(* Logix 5000 project; controller SmartManufacturingCell Emulate 5570 rev 33.11; software revision 33.03; part 4 of 5 *)
(* tags used below, declared in another part *)
   Production_CycleHealthy : BOOL;
   SequenceAtScan : DINT;
   StatisticsResetAccepted : BOOL;
   StatisticsResetONS : BOOL;
   Stats_ExitElapsed : REAL;
   Stats_HasPreviousExit : BOOL;
   Stats_RateElapsed : REAL;
   Stats_WindowCount : DINT;
   Conveyor_Flt_FailToStart : BOOL;   // Conveyor commanded but running feedback missing for 2 s Latched; clear cell, remove cause, then fresh Reset.
   Exit_Flt_DischargeTimeout : BOOL;   // Good or reject bottle departure not confirmed within 3 s Latched; clear cell, remove cause, then fresh Reset.
   Exit_Sts_GoodCompletePulse : BOOL;   // Exit Sts GoodCompletePulse
   Exit_Sts_RejectCompletePulse : BOOL;   // Exit Sts RejectCompletePulse
   Exit_Sts_State : DINT;   // 0 Empty; 10 Waiting; 20 Good discharge; 30 Extending; 40 Reject discharge; 50 Retracting; 60 Complete; 90 Faulted
   Filling_Flt_FillTimeout : BOOL;   // Fill completion not received within 4 s Latched; clear cell, remove cause, then fresh Reset.
   Filling_Flt_ValveFailToClose : BOOL;   // Fill valve did not close within 2 s Latched; clear cell, remove cause, then fresh Reset.
   Filling_Sts_ActiveFillTimeMs : DINT;   // Sampled fill duration for current bottle
   HMI_Cmd_Acknowledge : BOOL;   // Acknowledge alarm indication; does not reset faults
   HMI_Cmd_ClearCell : BOOL;   // Request removal of simulated bottles during fault recovery
   HMI_Cmd_ResetStatistics : BOOL;   // Clear production statistics only when Stopped and cell empty
   HMI_Cmd_Start : BOOL;   // Request automatic production start
   HMI_Cmd_Stop : BOOL;   // Request controlled production stop
   HMI_Sim_BottleMissingAtFill : BOOL;   // Suppress Fill photoeye while retaining simulated bottle presence. Simulation test only.
   HMI_Sim_ConveyorFailToStart : BOOL;   // Suppress conveyor running feedback. Simulation test only.
   HMI_Sim_FillFailToComplete : BOOL;   // Suppress simulated filling completion. Simulation test only.
   HMI_Sim_FillValveFailToClose : BOOL;   // Suppress fill valve closed feedback. Simulation test only.
   HMI_Sim_GoodDischargeJam : BOOL;   // Prevent good bottle departure. Simulation test only.
   HMI_Sim_IndexJam : BOOL;   // Prevent simulated index travel from completing. Simulation test only.
   HMI_Sim_IndexPositionMismatch : BOOL;   // Invert simulated Fill occupancy on transfer to test confirmation. Simulation test only.
   HMI_Sim_RejectDischargeJam : BOOL;   // Prevent rejected bottle departure. Simulation test only.
   HMI_Sim_RejectFailToExtend : BOOL;   // Suppress reject extended feedback. Simulation test only.
   HMI_Sim_RejectFailToRetract : BOOL;   // Suppress reject retracted feedback. Simulation test only.
   Inspection_Flt_Timeout : BOOL;   // Inspection did not finish within 3 s Latched; clear cell, remove cause, then fresh Reset.
   Production_Bottles : UDT_Bottle[4];
   Production_Flt_IndexConfirmTimeout : BOOL;   // Post-index positions not confirmed within 1 s Latched; clear cell, remove cause, then fresh Reset.
   Production_Flt_IndexInterlock : BOOL;   // Movement interlock lost during indexing Latched; clear cell, remove cause, then fresh Reset.
   Production_Flt_IndexTimeout : BOOL;   // Index completion not received within 3 s Latched; clear cell, remove cause, then fresh Reset.
   Production_Flt_InvalidConfiguration : BOOL;   // Fill or inspection time outside permitted limits Latched; clear cell, remove cause, then fresh Reset.
   Production_Flt_InvalidState : BOOL;   // Machine, sequence, station state, or mode combination invalid Latched; clear cell, remove cause, then fresh Reset.
   Production_Flt_StartupRecoveryRequired : BOOL;   // Restart found bottles or interrupted activity Latched; clear cell, remove cause, then fresh Reset.
   Production_Flt_TrackingMismatch : BOOL;   // Stationary bottle tracking and sensors disagree or processing history invalid Latched; clear cell, remove cause, then fr
   Production_Stats_FaultSeconds : REAL;   // FaultSeconds based on 20 ms scheduled executions; not a wall-clock historian.
   Production_Stats_GoodCount : DINT;   // Retained GoodCount; count only confirmed departures (recovery losses separate).
   Production_Stats_LastCycleSeconds : REAL;   // LastCycleSeconds based on 20 ms scheduled executions; not a wall-clock historian.
   Production_Stats_RatePerMinute : REAL;   // RatePerMinute based on 20 ms scheduled executions; not a wall-clock historian.
   Production_Stats_RecoveryLossCount : DINT;   // Retained RecoveryLossCount; count only confirmed departures (recovery losses separate).
   Production_Stats_RejectCount : DINT;   // Retained RejectCount; count only confirmed departures (recovery losses separate).
   Production_Stats_RunSeconds : REAL;   // RunSeconds based on 20 ms scheduled executions; not a wall-clock historian.
   Production_Stats_StoppedSeconds : REAL;   // StoppedSeconds based on 20 ms scheduled executions; not a wall-clock historian.
   Production_Stats_TotalCount : DINT;   // Retained TotalCount; count only confirmed departures (recovery losses separate).
   Production_Sts_ClearCellAccepted : BOOL;
   Production_Sts_CounterSaturated : BOOL;   // Production Sts CounterSaturated
   Production_Sts_IndexAllowed : BOOL;
   Production_Sts_IndexCommitted : BOOL;   // Bottle records transferred for the current confirmed index; cleared outside ConfirmPositions.
   Production_Sts_LoadAccepted : BOOL;
   Production_Sts_SequenceState : DINT;   // 0 = Idle 10 = ProcessStations 20 = Indexing 30 = ConfirmPositions
   Reject_Flt_FailToExtend : BOOL;   // Reject actuator did not extend within 2 s Latched; clear cell, remove cause, then fresh Reset.
   Reject_Flt_FailToRetract : BOOL;   // Reject actuator did not retract within 2 s Latched; clear cell, remove cause, then fresh Reset.
   Sim_In_ConveyorRunning : BOOL;   // Simulated conveyor movement feedback
   Sim_In_EntryPE : BOOL;   // Simulated bottle detected at entry
   Sim_In_ExitPE : BOOL;   // Simulated bottle detected at Reject/Exit position
   Sim_In_FillComplete : BOOL;   // Sim In FillComplete
   Sim_In_FillPE : BOOL;   // Simulated bottle detected at filling position
   Sim_In_FillValveClosed : BOOL;   // Simulated fill valve confirmed closed
   Sim_In_GoodExitPE : BOOL;   // Bottle detected passing through good discharge path
   Sim_In_IndexComplete : BOOL;   // Simulated conveyor completed one station-spacing movement
   Sim_In_InspectionPE : BOOL;   // Simulated bottle detected at inspection position
   Sim_In_RejectExitPE : BOOL;   // Bottle detected passing through reject discharge path
   Sim_In_RejectExtended : BOOL;   // Simulated reject actuator confirmed extended
   Sim_In_RejectRetracted : BOOL;   // Simulated reject actuator confirmed retracted
   Sim_Out_ConveyorRun : BOOL;   // Command simulated conveyor to run
   Sim_Out_FillValveOpen : BOOL;   // Command simulated fill valve to open
   Sim_Out_GoodDischargeRun : BOOL;   // Command simulated good-bottle discharge mechanism to run
   Sim_Out_RejectExtend : BOOL;   // Command simulated reject actuator to extend
   Sim_Sts_BottlesPresent : BOOL;   // Sim Sts BottlesPresent
   Sys_Sts_ActiveAlarmCount : DINT;   // Number of active latched faults
   Sys_Sts_AlarmUnacknowledged : BOOL;   // Sys Sts AlarmUnacknowledged
   Sys_Sts_AutoMode : BOOL;   // Auto mode accepted and active
   Sys_Sts_CellEmpty : BOOL;   // Sys Sts CellEmpty
   Sys_Sts_EquipmentHome : BOOL;   // Sys Sts EquipmentHome
   Sys_Sts_FirstFaultCode : DINT;   // Lowest active fault code; zero means none
   Sys_Sts_MachineState : DINT;   // 0 = Stopped 10 = Running 20 = Stopping 30 = Faulted
   Sys_Sts_ManualMode : BOOL;   // Manual mode accepted and active
   Sys_Sts_StartupReady : BOOL;   // Sys Sts StartupReady
(* Program_Production, continued *)

ROUTINE Production_Sequence   (* ladder *)
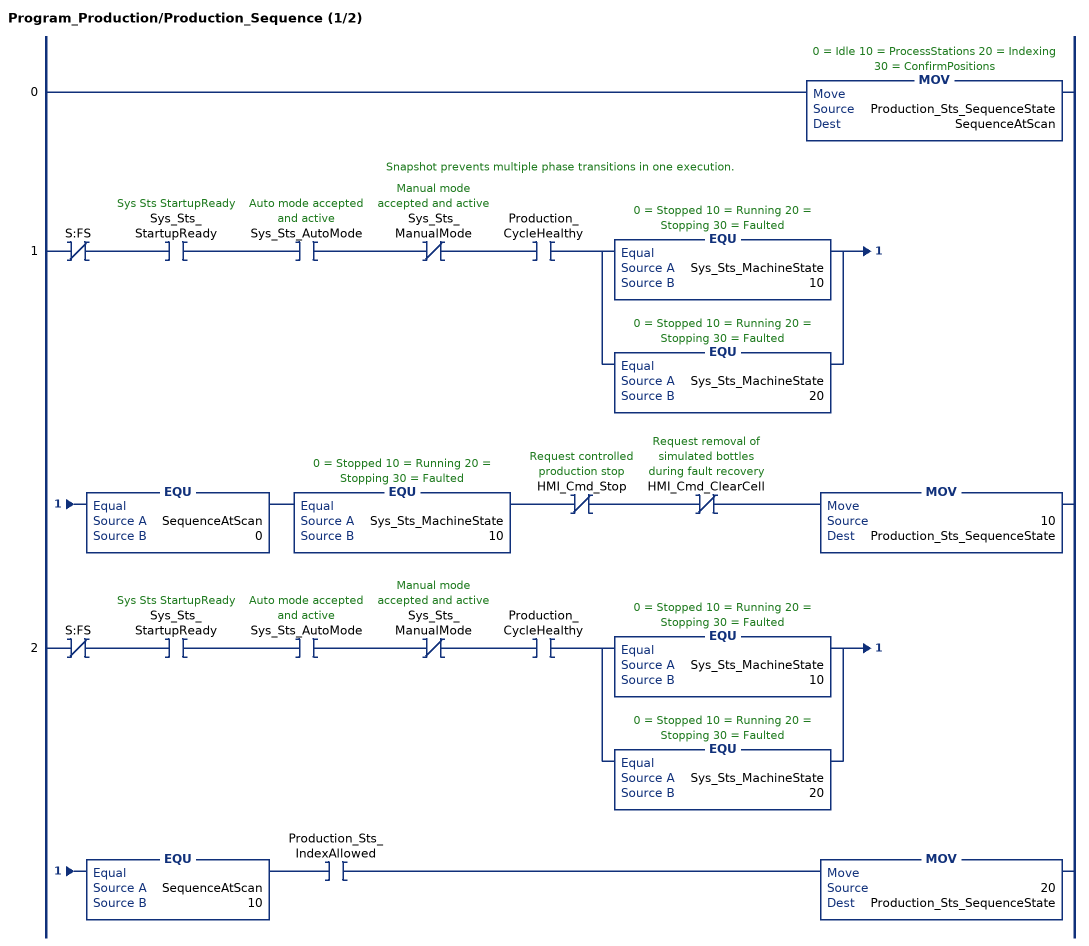
   0: MOV(Production_Sts_SequenceState,SequenceAtScan);
   // Snapshot prevents multiple phase transitions in one execution.
   1: XIO(S:FS)XIC(Sys_Sts_StartupReady)XIC(Sys_Sts_AutoMode)XIO(Sys_Sts_ManualMode)XIC(Production_CycleHealthy)[EQU(Sys_Sts_MachineState,10) ,EQU(Sys_Sts_MachineState,20) ]EQU(SequenceAtScan,0)EQU(Sys_Sts_MachineState,10)XIO(HMI_Cmd_Stop)XIO(HMI_Cmd_ClearCell)MOV(10,Production_Sts_SequenceState);
   2: XIO(S:FS)XIC(Sys_Sts_StartupReady)XIC(Sys_Sts_AutoMode)XIO(Sys_Sts_ManualMode)XIC(Production_CycleHealthy)[EQU(Sys_Sts_MachineState,10) ,EQU(Sys_Sts_MachineState,20) ]EQU(SequenceAtScan,10)XIC(Production_Sts_IndexAllowed)MOV(20,Production_Sts_SequenceState);
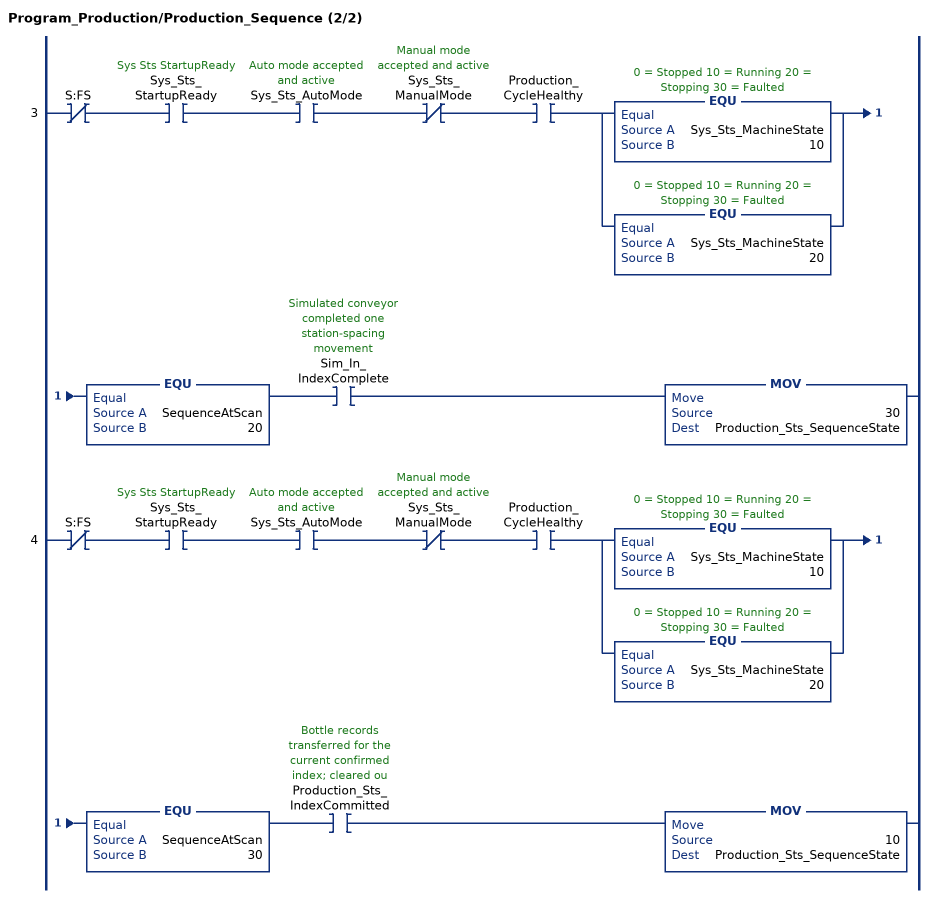
   3: XIO(S:FS)XIC(Sys_Sts_StartupReady)XIC(Sys_Sts_AutoMode)XIO(Sys_Sts_ManualMode)XIC(Production_CycleHealthy)[EQU(Sys_Sts_MachineState,10) ,EQU(Sys_Sts_MachineState,20) ]EQU(SequenceAtScan,20)XIC(Sim_In_IndexComplete)MOV(30,Production_Sts_SequenceState);
   4: XIO(S:FS)XIC(Sys_Sts_StartupReady)XIC(Sys_Sts_AutoMode)XIO(Sys_Sts_ManualMode)XIC(Production_CycleHealthy)[EQU(Sys_Sts_MachineState,10) ,EQU(Sys_Sts_MachineState,20) ]EQU(SequenceAtScan,30)XIC(Production_Sts_IndexCommitted)MOV(10,Production_Sts_SequenceState);
END_ROUTINE

ROUTINE Production_Statistics   (* structured text *)
   // One event per confirmed departure. Recovery clear losses are counted separately.
   IF Exit_Sts_GoodCompletePulse OR Exit_Sts_RejectCompletePulse THEN
       IF Production_Stats_TotalCount < 2147483647 THEN
           Production_Stats_TotalCount := Production_Stats_TotalCount + 1;
           IF Exit_Sts_GoodCompletePulse THEN
               Production_Stats_GoodCount := Production_Stats_GoodCount + 1;
           ELSE
               Production_Stats_RejectCount := Production_Stats_RejectCount + 1;
           END_IF;
       ELSE
           Production_Sts_CounterSaturated := 1;
       END_IF;
       IF Stats_HasPreviousExit THEN
           Production_Stats_LastCycleSeconds := Stats_ExitElapsed;
       END_IF;
       Stats_HasPreviousExit := 1;
       Stats_ExitElapsed := 0.0;
       Stats_WindowCount := Stats_WindowCount + 1;
       Production_Bottles[3].Occupied := 0;
       Production_Bottles[3].FillComplete := 0;
       Production_Bottles[3].InspectionComplete := 0;
       Production_Bottles[3].RejectRequired := 0;
   END_IF;
   IF (Sys_Sts_MachineState = 10) OR (Sys_Sts_MachineState = 20) THEN
       Production_Stats_RunSeconds := Production_Stats_RunSeconds + 0.02;
       Stats_ExitElapsed := Stats_ExitElapsed + 0.02;
   ELSIF Sys_Sts_MachineState = 30 THEN
       Production_Stats_FaultSeconds := Production_Stats_FaultSeconds + 0.02;
   ELSE
       Production_Stats_StoppedSeconds := Production_Stats_StoppedSeconds + 0.02;
   END_IF;
   Stats_RateElapsed := Stats_RateElapsed + 0.02;
   IF Stats_RateElapsed >= 60.0 THEN
       Production_Stats_RatePerMinute := Stats_WindowCount * 60.0 / Stats_RateElapsed;
       Stats_RateElapsed := 0.0;
       Stats_WindowCount := 0;
   END_IF;
   IF S:FS THEN
       Stats_ExitElapsed := 0.0;
       Stats_HasPreviousExit := 0;
       Stats_RateElapsed := 0.0;
       Stats_WindowCount := 0;
       Production_Stats_RatePerMinute := 0.0;
   END_IF;
   IF StatisticsResetAccepted THEN
       Production_Stats_TotalCount := 0;
       Production_Stats_GoodCount := 0;
       Production_Stats_RejectCount := 0;
       Production_Stats_RecoveryLossCount := 0;
       Production_Stats_RunSeconds := 0.0;
       Production_Stats_StoppedSeconds := 0.0;
       Production_Stats_FaultSeconds := 0.0;
       Production_Stats_LastCycleSeconds := 0.0;
       Production_Stats_RatePerMinute := 0.0;
       Production_Sts_CounterSaturated := 0;
       Stats_ExitElapsed := 0.0;
       Stats_HasPreviousExit := 0;
       Stats_RateElapsed := 0.0;
       Stats_WindowCount := 0;
   END_IF;
END_ROUTINE

ROUTINE Statistics_Reset   (* ladder *)
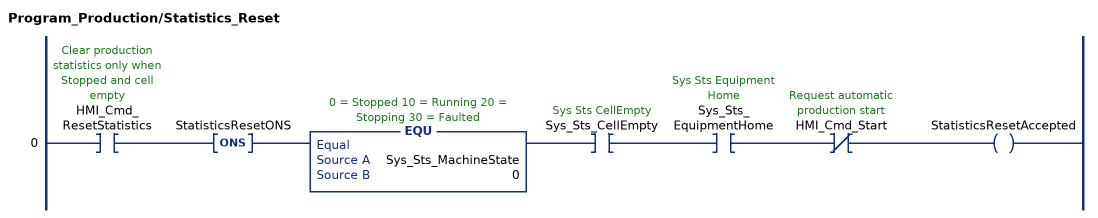
   0: XIC(HMI_Cmd_ResetStatistics)ONS(StatisticsResetONS)EQU(Sys_Sts_MachineState,0)XIC(Sys_Sts_CellEmpty)XIC(Sys_Sts_EquipmentHome)XIO(HMI_Cmd_Start)OTE(StatisticsResetAccepted);
END_ROUTINE
END_PROGRAM

PROGRAM Program_Simulation   (* main routine Main_Routine *)
VAR
   ConveyorStartDelay : TIMER := (PRE := 200); {access None}   // Non-retentive timer; preset in milliseconds.
   FillProcessDelay : TIMER := (PRE := 1500); {access None}   // Non-retentive timer; preset in milliseconds.
   FillValveCloseDelay : TIMER := (PRE := 150); {access None}   // Non-retentive timer; preset in milliseconds.
   GoodDischargeDelay : TIMER := (PRE := 700); {access None}   // Non-retentive timer; preset in milliseconds.
   GoodTransferONS : BOOL; {access None}
   GoodTransferPulse : BOOL; {access None}
   IndexTransferONS : BOOL; {access None}
   IndexTransferPulse : BOOL; {access None}
   IndexTravelDelay : TIMER := (PRE := 1000); {access None}   // Non-retentive timer; preset in milliseconds.
   RejectDischargeDelay : TIMER := (PRE := 500); {access None}   // Non-retentive timer; preset in milliseconds.
   RejectExtendDelay : TIMER := (PRE := 200); {access None}   // Non-retentive timer; preset in milliseconds.
   RejectRetractDelay : TIMER := (PRE := 200); {access None}   // Non-retentive timer; preset in milliseconds.
   RejectTransferONS : BOOL; {access None}
   RejectTransferPulse : BOOL; {access None}
   Sim_EntryOccupied : BOOL; {access None}   // Simulated physical bottle presence at Entry.
   Sim_ExitOccupied : BOOL; {access None}
   Sim_FillOccupied : BOOL; {access None}
   Sim_InspectionOccupied : BOOL; {access None}
END_VAR

ROUTINE Bottle_Simulation   (* ladder *)
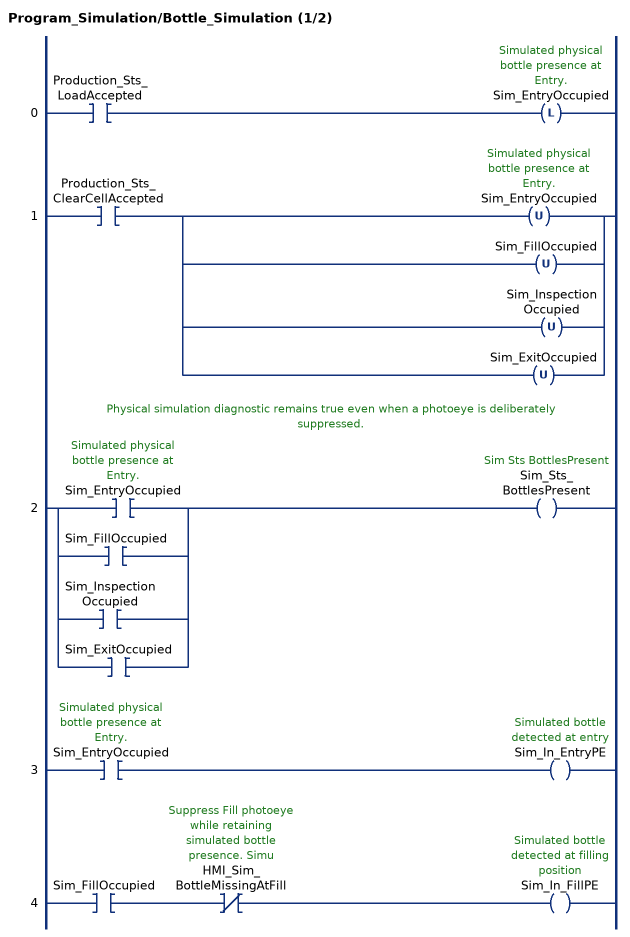
   0: XIC(Production_Sts_LoadAccepted)OTL(Sim_EntryOccupied);
   1: XIC(Production_Sts_ClearCellAccepted)[OTU(Sim_EntryOccupied) ,OTU(Sim_FillOccupied) ,OTU(Sim_InspectionOccupied) ,OTU(Sim_ExitOccupied) ];
   // Physical simulation diagnostic remains true even when a photoeye is deliberately suppressed.
   2: [XIC(Sim_EntryOccupied) ,XIC(Sim_FillOccupied) ,XIC(Sim_InspectionOccupied) ,XIC(Sim_ExitOccupied) ]OTE(Sim_Sts_BottlesPresent);
   3: XIC(Sim_EntryOccupied)OTE(Sim_In_EntryPE);
   4: XIC(Sim_FillOccupied)XIO(HMI_Sim_BottleMissingAtFill)OTE(Sim_In_FillPE);
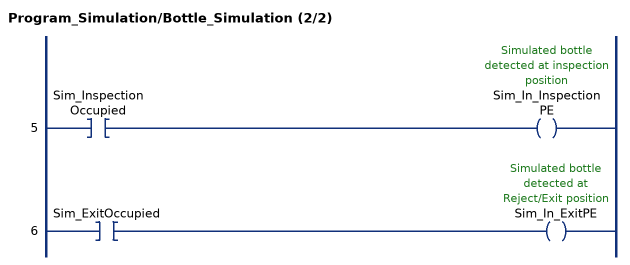
   5: XIC(Sim_InspectionOccupied)OTE(Sim_In_InspectionPE);
   6: XIC(Sim_ExitOccupied)OTE(Sim_In_ExitPE);
END_ROUTINE

ROUTINE Conveyor_Simulation   (* ladder *)
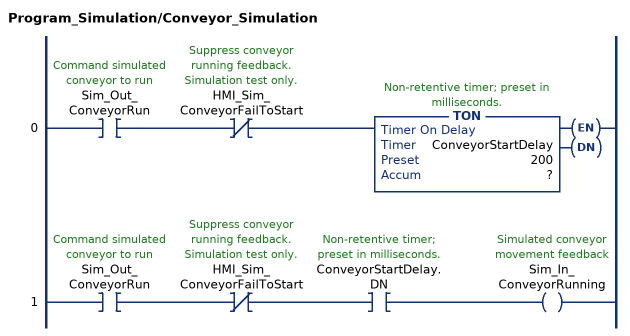
   0: XIC(Sim_Out_ConveyorRun)XIO(HMI_Sim_ConveyorFailToStart)TON(ConveyorStartDelay,?,?);
   1: XIC(Sim_Out_ConveyorRun)XIO(HMI_Sim_ConveyorFailToStart)XIC(ConveyorStartDelay.DN)OTE(Sim_In_ConveyorRunning);
END_ROUTINE

ROUTINE Exit_Simulation   (* ladder *)
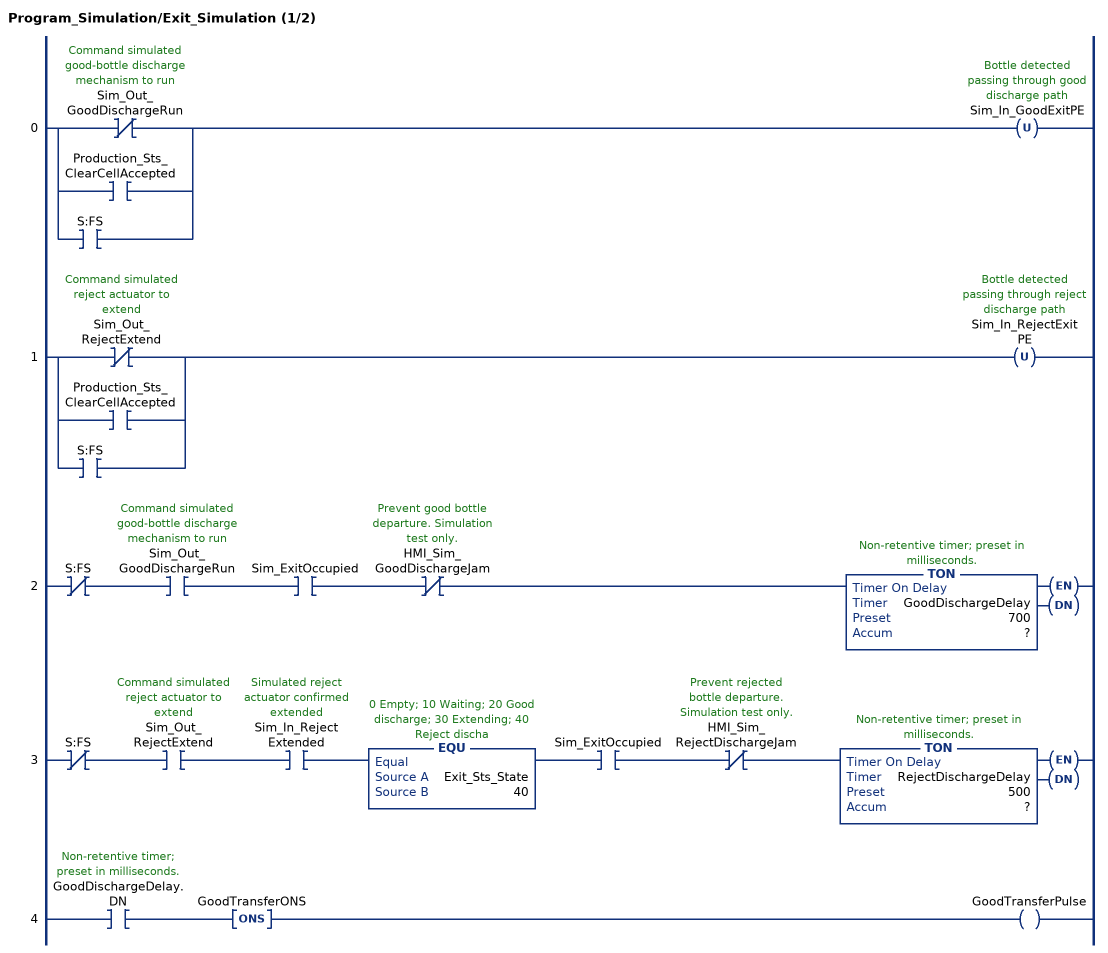
   0: [XIO(Sim_Out_GoodDischargeRun) ,XIC(Production_Sts_ClearCellAccepted) ,XIC(S:FS) ]OTU(Sim_In_GoodExitPE);
   1: [XIO(Sim_Out_RejectExtend) ,XIC(Production_Sts_ClearCellAccepted) ,XIC(S:FS) ]OTU(Sim_In_RejectExitPE);
   2: XIO(S:FS)XIC(Sim_Out_GoodDischargeRun)XIC(Sim_ExitOccupied)XIO(HMI_Sim_GoodDischargeJam)TON(GoodDischargeDelay,?,?);
   3: XIO(S:FS)XIC(Sim_Out_RejectExtend)XIC(Sim_In_RejectExtended)EQU(Exit_Sts_State,40)XIC(Sim_ExitOccupied)XIO(HMI_Sim_RejectDischargeJam)TON(RejectDischargeDelay,?,?);
   4: XIC(GoodDischargeDelay.DN)ONS(GoodTransferONS)OTE(GoodTransferPulse);
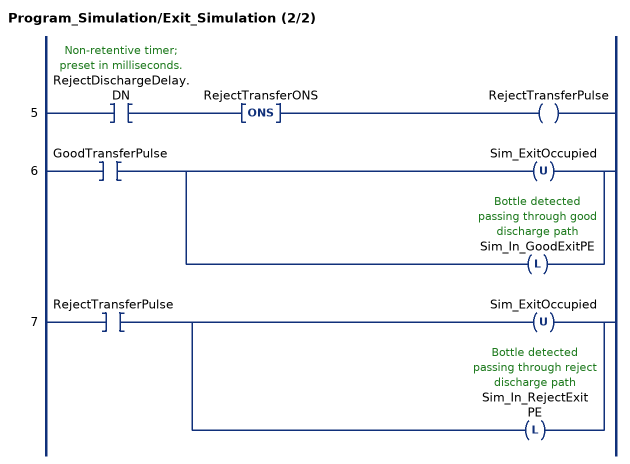
   5: XIC(RejectDischargeDelay.DN)ONS(RejectTransferONS)OTE(RejectTransferPulse);
   6: XIC(GoodTransferPulse)[OTU(Sim_ExitOccupied) ,OTL(Sim_In_GoodExitPE) ];
   7: XIC(RejectTransferPulse)[OTU(Sim_ExitOccupied) ,OTL(Sim_In_RejectExitPE) ];
END_ROUTINE

ROUTINE Filling_Simulation   (* ladder *)
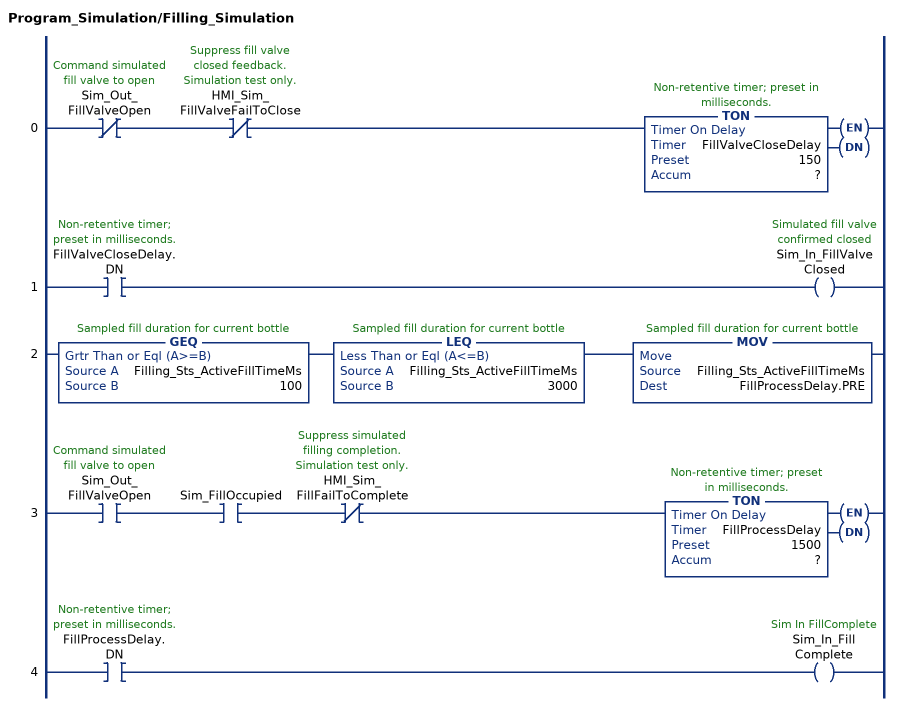
   0: XIO(Sim_Out_FillValveOpen)XIO(HMI_Sim_FillValveFailToClose)TON(FillValveCloseDelay,?,?);
   1: XIC(FillValveCloseDelay.DN)OTE(Sim_In_FillValveClosed);
   2: GEQ(Filling_Sts_ActiveFillTimeMs,100)LEQ(Filling_Sts_ActiveFillTimeMs,3000)MOV(Filling_Sts_ActiveFillTimeMs,FillProcessDelay.PRE);
   3: XIC(Sim_Out_FillValveOpen)XIC(Sim_FillOccupied)XIO(HMI_Sim_FillFailToComplete)TON(FillProcessDelay,?,?);
   4: XIC(FillProcessDelay.DN)OTE(Sim_In_FillComplete);
END_ROUTINE

ROUTINE Index_Simulation   (* ladder *)
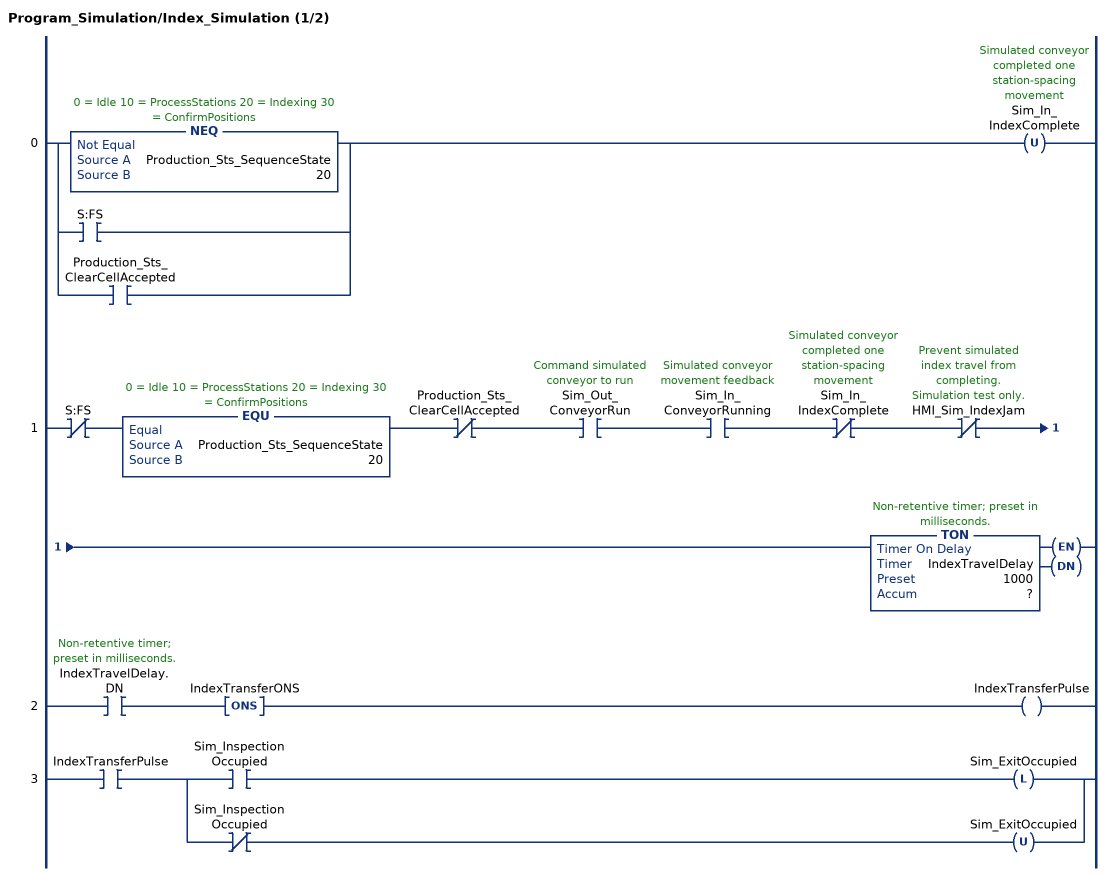
   0: [NEQ(Production_Sts_SequenceState,20) ,XIC(S:FS) ,XIC(Production_Sts_ClearCellAccepted) ]OTU(Sim_In_IndexComplete);
   1: XIO(S:FS)EQU(Production_Sts_SequenceState,20)XIO(Production_Sts_ClearCellAccepted)XIC(Sim_Out_ConveyorRun)XIC(Sim_In_ConveyorRunning)XIO(Sim_In_IndexComplete)XIO(HMI_Sim_IndexJam)TON(IndexTravelDelay,?,?);
   2: XIC(IndexTravelDelay.DN)ONS(IndexTransferONS)OTE(IndexTransferPulse);
   3: XIC(IndexTransferPulse)[XIC(Sim_InspectionOccupied) OTL(Sim_ExitOccupied) ,XIO(Sim_InspectionOccupied) OTU(Sim_ExitOccupied) ];
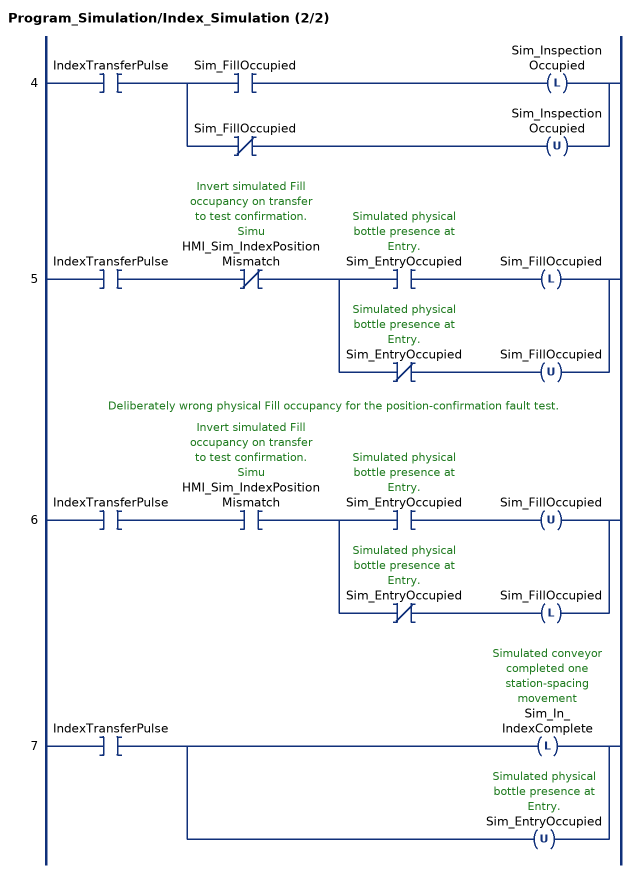
   4: XIC(IndexTransferPulse)[XIC(Sim_FillOccupied) OTL(Sim_InspectionOccupied) ,XIO(Sim_FillOccupied) OTU(Sim_InspectionOccupied) ];
   5: XIC(IndexTransferPulse)XIO(HMI_Sim_IndexPositionMismatch)[XIC(Sim_EntryOccupied) OTL(Sim_FillOccupied) ,XIO(Sim_EntryOccupied) OTU(Sim_FillOccupied) ];
   // Deliberately wrong physical Fill occupancy for the position-confirmation fault test.
   6: XIC(IndexTransferPulse)XIC(HMI_Sim_IndexPositionMismatch)[XIC(Sim_EntryOccupied) OTU(Sim_FillOccupied) ,XIO(Sim_EntryOccupied) OTL(Sim_FillOccupied) ];
   7: XIC(IndexTransferPulse)[OTL(Sim_In_IndexComplete) ,OTU(Sim_EntryOccupied) ];
END_ROUTINE

ROUTINE Main_Routine   (* ladder *)
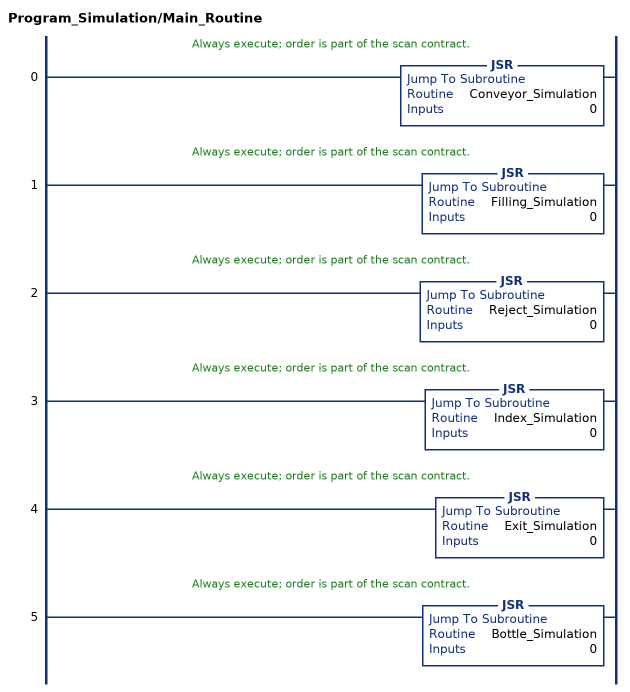
   // Always execute; order is part of the scan contract.
   0: JSR(Conveyor_Simulation,0);
   // Always execute; order is part of the scan contract.
   1: JSR(Filling_Simulation,0);
   // Always execute; order is part of the scan contract.
   2: JSR(Reject_Simulation,0);
   // Always execute; order is part of the scan contract.
   3: JSR(Index_Simulation,0);
   // Always execute; order is part of the scan contract.
   4: JSR(Exit_Simulation,0);
   // Always execute; order is part of the scan contract.
   5: JSR(Bottle_Simulation,0);
END_ROUTINE

ROUTINE Reject_Simulation   (* ladder *)
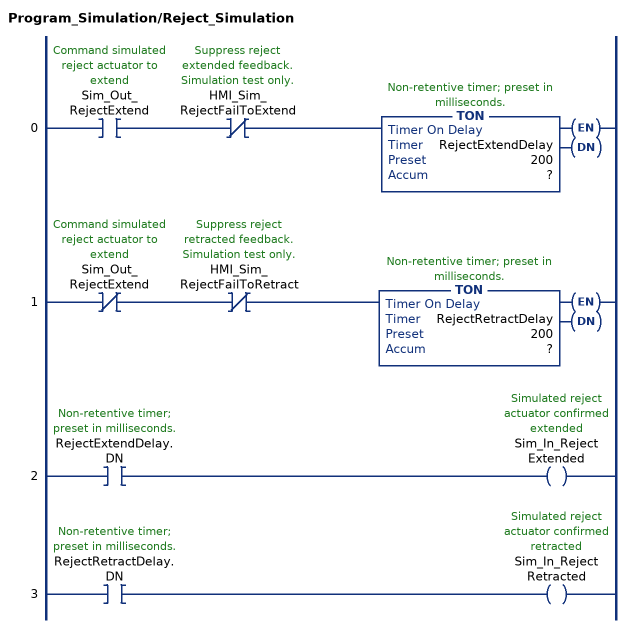
   0: XIC(Sim_Out_RejectExtend)XIO(HMI_Sim_RejectFailToExtend)TON(RejectExtendDelay,?,?);
   1: XIO(Sim_Out_RejectExtend)XIO(HMI_Sim_RejectFailToRetract)TON(RejectRetractDelay,?,?);
   2: XIC(RejectExtendDelay.DN)OTE(Sim_In_RejectExtended);
   3: XIC(RejectRetractDelay.DN)OTE(Sim_In_RejectRetracted);
END_ROUTINE
END_PROGRAM

PROGRAM Program_System   (* main routine MainRoutine *)
// Machine mode, startup, controlled stop, and overall fault coordination.
VAR
   AlarmAckONS : BOOL; {access None}
   AlarmEdge101 : BOOL; {access None}
   AlarmEdge201 : BOOL; {access None}
   AlarmEdge202 : BOOL; {access None}
   AlarmEdge301 : BOOL; {access None}
   AlarmEdge401 : BOOL; {access None}
   AlarmEdge402 : BOOL; {access None}
   AlarmEdge403 : BOOL; {access None}
   AlarmEdge501 : BOOL; {access None}
   AlarmEdge502 : BOOL; {access None}
   AlarmEdge503 : BOOL; {access None}
   AlarmEdge504 : BOOL; {access None}
   AlarmEdge505 : BOOL; {access None}
   AlarmEdge506 : BOOL; {access None}
   AlarmEdge507 : BOOL; {access None}
   AutoRequestONS : BOOL; {access Read Only}
   ConfigurationValid : BOOL; {access None}
   ManualRequestONS : BOOL; {access Read Only}
   ModeChangeAllowed : BOOL; {access Read Only}
   Recovery_CommandsReleased : BOOL; {access None}
   Recovery_PhaseClear : BOOL; {access None}
   Recovery_SensorsClear : BOOL; {access None}
   Recovery_TrackingClear : BOOL; {access None}
   Start_CommandsReleased : BOOL; {access None}
   Start_EquipmentReady : BOOL; {access None}
   StartRequestONS : BOOL; {access None}
   Startup_CheckPending : BOOL; {access None}
END_VAR

ROUTINE Alarm_Control   (* ladder *)
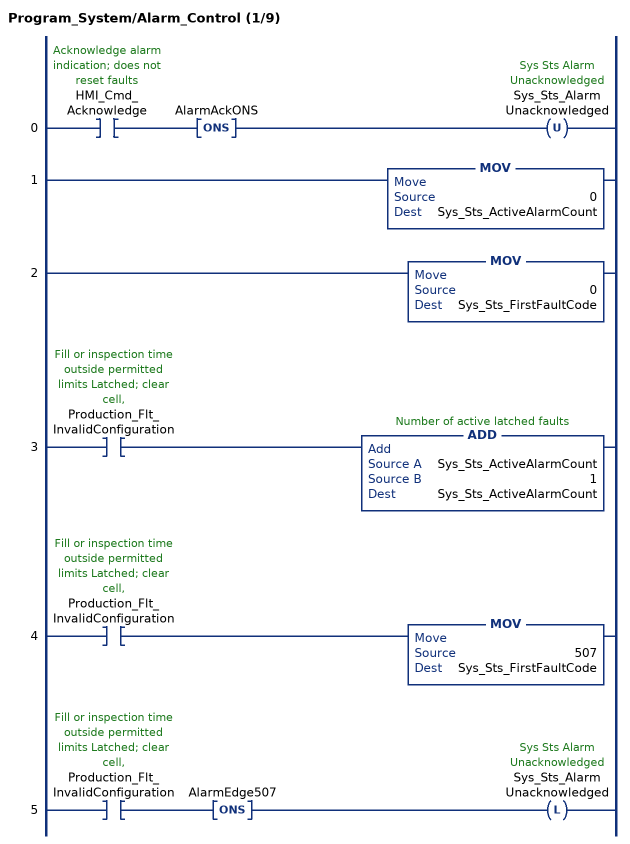
   0: XIC(HMI_Cmd_Acknowledge)ONS(AlarmAckONS)OTU(Sys_Sts_AlarmUnacknowledged);
   1: MOV(0,Sys_Sts_ActiveAlarmCount);
   2: MOV(0,Sys_Sts_FirstFaultCode);
   3: XIC(Production_Flt_InvalidConfiguration)ADD(Sys_Sts_ActiveAlarmCount,1,Sys_Sts_ActiveAlarmCount);
   4: XIC(Production_Flt_InvalidConfiguration)MOV(507,Sys_Sts_FirstFaultCode);
   5: XIC(Production_Flt_InvalidConfiguration)ONS(AlarmEdge507)OTL(Sys_Sts_AlarmUnacknowledged);
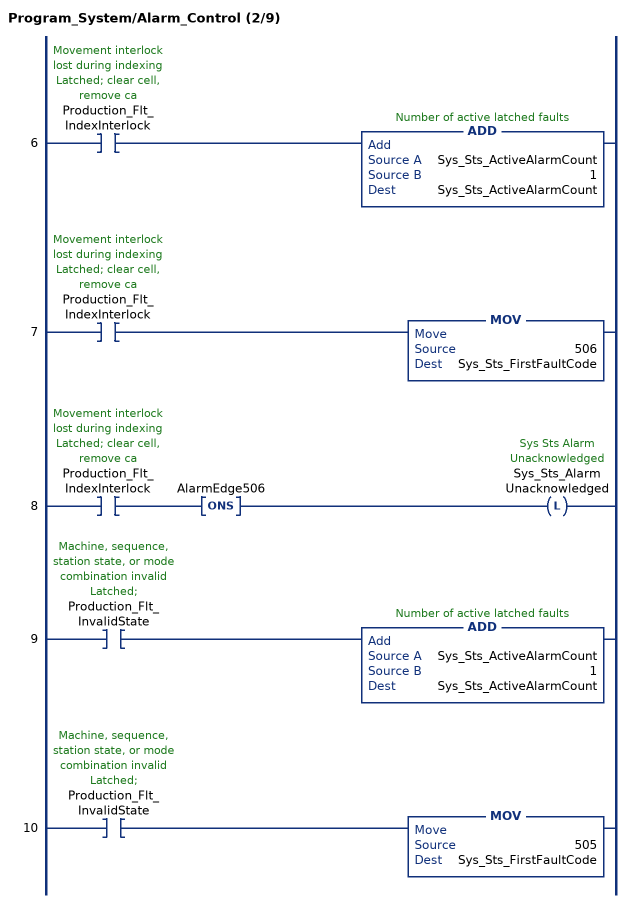
   6: XIC(Production_Flt_IndexInterlock)ADD(Sys_Sts_ActiveAlarmCount,1,Sys_Sts_ActiveAlarmCount);
   7: XIC(Production_Flt_IndexInterlock)MOV(506,Sys_Sts_FirstFaultCode);
   8: XIC(Production_Flt_IndexInterlock)ONS(AlarmEdge506)OTL(Sys_Sts_AlarmUnacknowledged);
   9: XIC(Production_Flt_InvalidState)ADD(Sys_Sts_ActiveAlarmCount,1,Sys_Sts_ActiveAlarmCount);
   10: XIC(Production_Flt_InvalidState)MOV(505,Sys_Sts_FirstFaultCode);
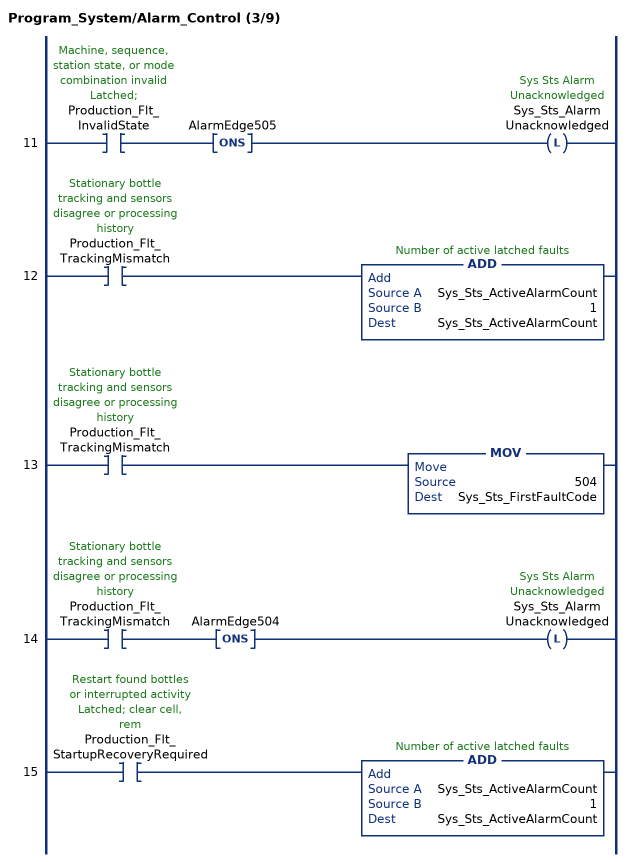
   11: XIC(Production_Flt_InvalidState)ONS(AlarmEdge505)OTL(Sys_Sts_AlarmUnacknowledged);
   12: XIC(Production_Flt_TrackingMismatch)ADD(Sys_Sts_ActiveAlarmCount,1,Sys_Sts_ActiveAlarmCount);
   13: XIC(Production_Flt_TrackingMismatch)MOV(504,Sys_Sts_FirstFaultCode);
   14: XIC(Production_Flt_TrackingMismatch)ONS(AlarmEdge504)OTL(Sys_Sts_AlarmUnacknowledged);
   15: XIC(Production_Flt_StartupRecoveryRequired)ADD(Sys_Sts_ActiveAlarmCount,1,Sys_Sts_ActiveAlarmCount);
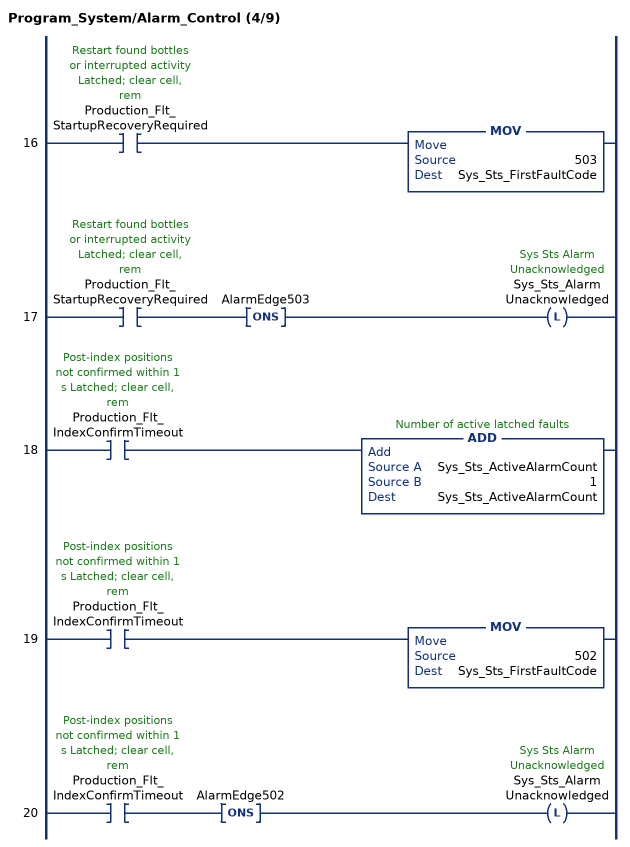
   16: XIC(Production_Flt_StartupRecoveryRequired)MOV(503,Sys_Sts_FirstFaultCode);
   17: XIC(Production_Flt_StartupRecoveryRequired)ONS(AlarmEdge503)OTL(Sys_Sts_AlarmUnacknowledged);
   18: XIC(Production_Flt_IndexConfirmTimeout)ADD(Sys_Sts_ActiveAlarmCount,1,Sys_Sts_ActiveAlarmCount);
   19: XIC(Production_Flt_IndexConfirmTimeout)MOV(502,Sys_Sts_FirstFaultCode);
   20: XIC(Production_Flt_IndexConfirmTimeout)ONS(AlarmEdge502)OTL(Sys_Sts_AlarmUnacknowledged);
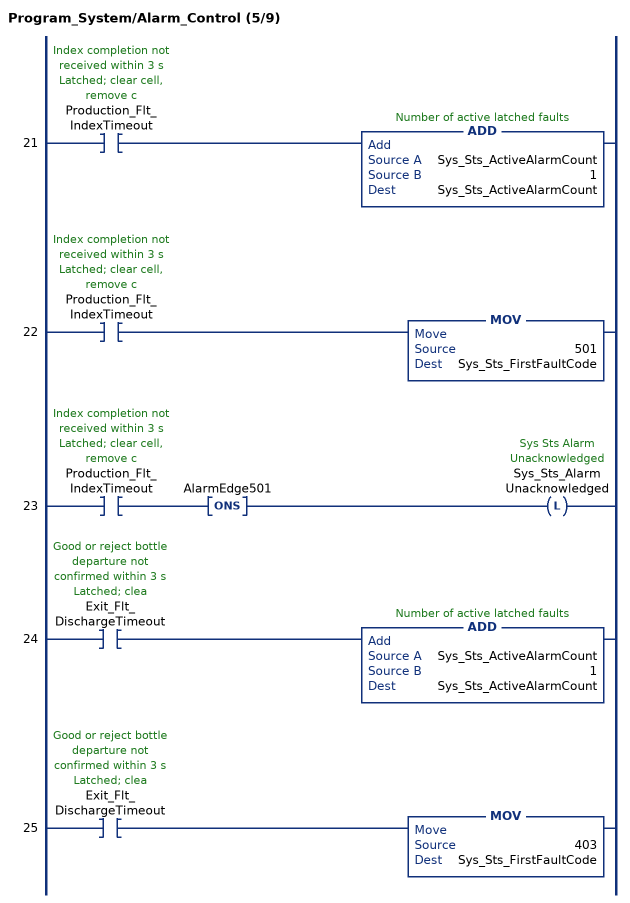
   21: XIC(Production_Flt_IndexTimeout)ADD(Sys_Sts_ActiveAlarmCount,1,Sys_Sts_ActiveAlarmCount);
   22: XIC(Production_Flt_IndexTimeout)MOV(501,Sys_Sts_FirstFaultCode);
   23: XIC(Production_Flt_IndexTimeout)ONS(AlarmEdge501)OTL(Sys_Sts_AlarmUnacknowledged);
   24: XIC(Exit_Flt_DischargeTimeout)ADD(Sys_Sts_ActiveAlarmCount,1,Sys_Sts_ActiveAlarmCount);
   25: XIC(Exit_Flt_DischargeTimeout)MOV(403,Sys_Sts_FirstFaultCode);
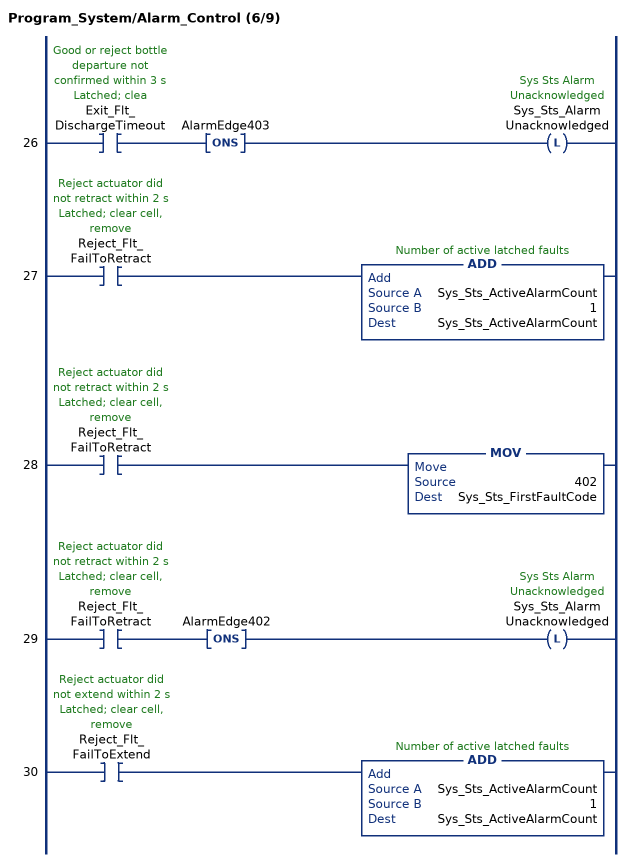
   26: XIC(Exit_Flt_DischargeTimeout)ONS(AlarmEdge403)OTL(Sys_Sts_AlarmUnacknowledged);
   27: XIC(Reject_Flt_FailToRetract)ADD(Sys_Sts_ActiveAlarmCount,1,Sys_Sts_ActiveAlarmCount);
   28: XIC(Reject_Flt_FailToRetract)MOV(402,Sys_Sts_FirstFaultCode);
   29: XIC(Reject_Flt_FailToRetract)ONS(AlarmEdge402)OTL(Sys_Sts_AlarmUnacknowledged);
   30: XIC(Reject_Flt_FailToExtend)ADD(Sys_Sts_ActiveAlarmCount,1,Sys_Sts_ActiveAlarmCount);
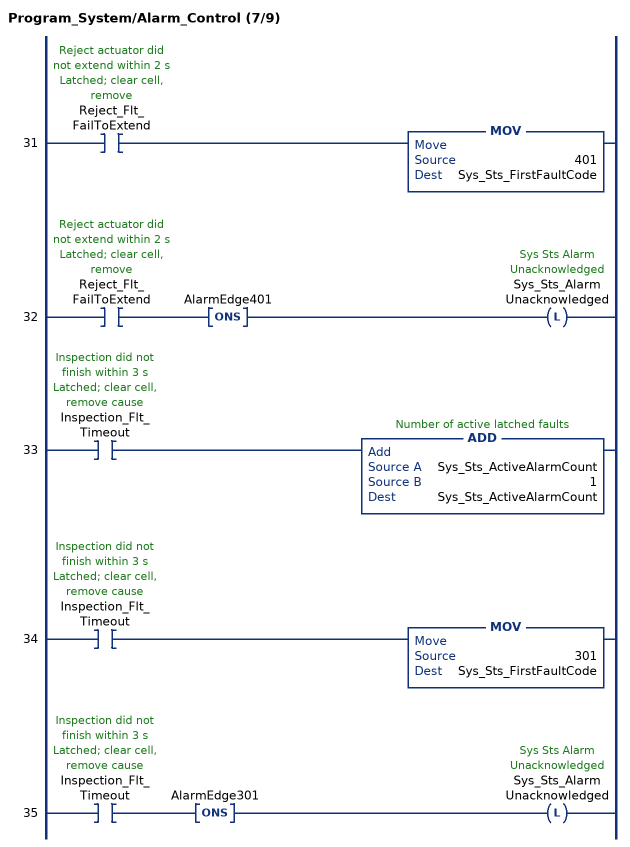
   31: XIC(Reject_Flt_FailToExtend)MOV(401,Sys_Sts_FirstFaultCode);
   32: XIC(Reject_Flt_FailToExtend)ONS(AlarmEdge401)OTL(Sys_Sts_AlarmUnacknowledged);
   33: XIC(Inspection_Flt_Timeout)ADD(Sys_Sts_ActiveAlarmCount,1,Sys_Sts_ActiveAlarmCount);
   34: XIC(Inspection_Flt_Timeout)MOV(301,Sys_Sts_FirstFaultCode);
   35: XIC(Inspection_Flt_Timeout)ONS(AlarmEdge301)OTL(Sys_Sts_AlarmUnacknowledged);
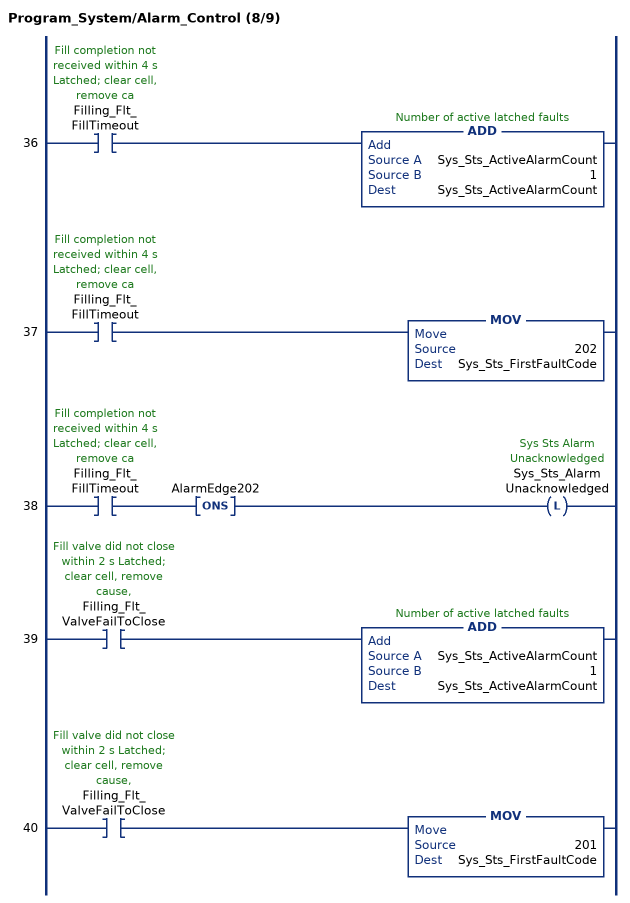
   36: XIC(Filling_Flt_FillTimeout)ADD(Sys_Sts_ActiveAlarmCount,1,Sys_Sts_ActiveAlarmCount);
   37: XIC(Filling_Flt_FillTimeout)MOV(202,Sys_Sts_FirstFaultCode);
   38: XIC(Filling_Flt_FillTimeout)ONS(AlarmEdge202)OTL(Sys_Sts_AlarmUnacknowledged);
   39: XIC(Filling_Flt_ValveFailToClose)ADD(Sys_Sts_ActiveAlarmCount,1,Sys_Sts_ActiveAlarmCount);
   40: XIC(Filling_Flt_ValveFailToClose)MOV(201,Sys_Sts_FirstFaultCode);
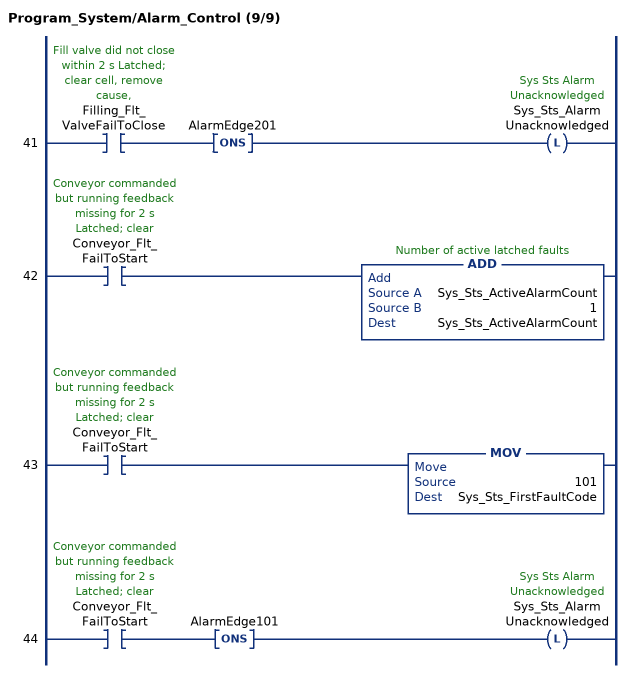
   41: XIC(Filling_Flt_ValveFailToClose)ONS(AlarmEdge201)OTL(Sys_Sts_AlarmUnacknowledged);
   42: XIC(Conveyor_Flt_FailToStart)ADD(Sys_Sts_ActiveAlarmCount,1,Sys_Sts_ActiveAlarmCount);
   43: XIC(Conveyor_Flt_FailToStart)MOV(101,Sys_Sts_FirstFaultCode);
   44: XIC(Conveyor_Flt_FailToStart)ONS(AlarmEdge101)OTL(Sys_Sts_AlarmUnacknowledged);
END_ROUTINE
